(* IEC 61131-3 sources: RootPLC/conformance/cases/motion, 8 files *)

(* ---- ok_abort_and_relative.st ---- *)
(* spec: [motion.abort] [motion.move.relative]
   expect: ok
   libraries: RootMotion *)
TEST new_command_takes_control_without_a_jump
VAR
    ax : AXIS_REF;
    pw : MC_Power;
    m1 : MC_MoveAbsolute;
    m2 : MC_MoveRelative;
    i : INT;
    startPos : LREAL;
    vBefore : LREAL;
END_VAR
ax.CycleTime := 0.01;
pw(Enable := TRUE, Axis := ax);
FOR i := 1 TO 20 DO
    m1(Execute := TRUE, Position := 100.0, Velocity := 50.0, Acceleration := 100.0, Deceleration := 100.0, Axis := ax);
    RP_VirtualAxis(Axis := ax);
END_FOR;
startPos := ax.Position;
vBefore := ax.Velocity;
m2(Execute := TRUE, Distance := -5.0, Velocity := 50.0, Acceleration := 100.0, Deceleration := 100.0, Axis := ax);
m1(Execute := TRUE, Position := 100.0, Velocity := 50.0, Acceleration := 100.0, Deceleration := 100.0, Axis := ax);
ASSERT_TRUE(m1.CommandAborted);
ASSERT_FALSE(m1.Busy);
RP_VirtualAxis(Axis := ax);
ASSERT_TRUE(ABS(ax.Velocity - vBefore) <= 1.000001);
FOR i := 1 TO 300 DO
    m2(Execute := TRUE, Distance := -5.0, Velocity := 50.0, Acceleration := 100.0, Deceleration := 100.0, Axis := ax);
    RP_VirtualAxis(Axis := ax);
END_FOR;
ASSERT_TRUE(m2.Done);
ASSERT_TRUE(ABS(ax.Position - (startPos - 5.0)) < 0.000001);
END_TEST

(* ---- ok_errors_and_execute.st ---- *)
(* spec: [motion.errors] [motion.execute] [motion.power]
   expect: ok
   libraries: RootMotion *)
TEST command_on_unpowered_axis
VAR
    ax : AXIS_REF;
    mv : MC_MoveAbsolute;
END_VAR
mv(Execute := TRUE, Position := 10.0, Velocity := 5.0, Acceleration := 10.0, Deceleration := 10.0, Axis := ax);
ASSERT_TRUE(mv.Error);
ASSERT_EQ(UDINT#1, mv.ErrorID);
ASSERT_TRUE(ax.State = MC_AXIS_STATE#Disabled);
END_TEST

TEST invalid_parameter
VAR
    ax : AXIS_REF;
    pw : MC_Power;
    mv : MC_MoveAbsolute;
END_VAR
pw(Enable := TRUE, Axis := ax);
mv(Execute := TRUE, Position := 10.0, Velocity := 0.0, Acceleration := 10.0, Deceleration := 10.0, Axis := ax);
ASSERT_TRUE(mv.Error);
ASSERT_EQ(UDINT#3, mv.ErrorID);
ASSERT_TRUE(ax.State = MC_AXIS_STATE#Standstill);
END_TEST

TEST result_shows_one_call_after_execute_falls
VAR
    ax : AXIS_REF;
    pw : MC_Power;
    mv : MC_MoveAbsolute;
    i : INT;
END_VAR
ax.CycleTime := 0.1;
pw(Enable := TRUE, Axis := ax);
mv(Execute := TRUE, Position := 1.0, Velocity := 10.0, Acceleration := 100.0, Deceleration := 100.0, Axis := ax);
FOR i := 1 TO 20 DO
    mv(Execute := FALSE, Position := 1.0, Velocity := 10.0, Acceleration := 100.0, Deceleration := 100.0, Axis := ax);
    RP_VirtualAxis(Axis := ax);
    IF mv.Done THEN
        EXIT;
    END_IF;
END_FOR;
ASSERT_TRUE(mv.Done);
ASSERT_TRUE(ABS(ax.Position - 1.0) < 0.000001);
mv(Execute := FALSE, Position := 1.0, Velocity := 10.0, Acceleration := 100.0, Deceleration := 100.0, Axis := ax);
ASSERT_FALSE(mv.Done);
END_TEST

(* ---- ok_home.st ---- *)
(* spec: [motion.home] [motion.errors]
   expect: ok
   libraries: RootMotion *)
TEST home_sets_position
VAR
    ax : AXIS_REF;
    pw : MC_Power;
    hm : MC_Home;
END_VAR
hm(Execute := TRUE, Position := 0.0, Axis := ax);
ASSERT_TRUE(hm.Error);
ASSERT_EQ(UDINT#1, hm.ErrorID);
hm(Execute := FALSE, Position := 0.0, Axis := ax);
pw(Enable := TRUE, Axis := ax);
hm(Execute := TRUE, Position := 12.5, Axis := ax);
ASSERT_TRUE(hm.Done);
ASSERT_TRUE(ax.Homed);
ASSERT_TRUE(ABS(ax.Position - 12.5) < 0.000001);
ASSERT_TRUE(ax.State = MC_AXIS_STATE#Standstill);
END_TEST

(* ---- ok_limits_reset_stop.st ---- *)
(* spec: [motion.limits] [motion.reset] [motion.stop] [motion.errors]
   expect: ok
   libraries: RootMotion *)
TEST limit_error_reset_then_stop
VAR
    ax : AXIS_REF;
    pw : MC_Power;
    mvv : MC_MoveVelocity;
    mv : MC_MoveAbsolute;
    st : MC_Stop;
    rs : MC_Reset;
    i : INT;
END_VAR
ax.CycleTime := 0.01;
ax.LimitsEnabled := TRUE;
ax.PositiveLimit := 50.0;
ax.NegativeLimit := -50.0;
pw(Enable := TRUE, Axis := ax);
FOR i := 1 TO 600 DO
    mvv(Execute := TRUE, Velocity := 20.0, Acceleration := 100.0, Deceleration := 100.0, Axis := ax);
    RP_VirtualAxis(Axis := ax);
END_FOR;
mvv(Execute := TRUE, Velocity := 20.0, Acceleration := 100.0, Deceleration := 100.0, Axis := ax);
ASSERT_TRUE(ax.State = MC_AXIS_STATE#ErrorStop);
ASSERT_TRUE(mvv.Error);
ASSERT_EQ(UDINT#4, mvv.ErrorID);
ASSERT_TRUE(ABS(ax.Position - 50.0) < 0.000001);
ASSERT_TRUE(ABS(ax.Velocity) < 0.000001);
mv(Execute := TRUE, Position := 0.0, Velocity := 10.0, Acceleration := 100.0, Deceleration := 100.0, Axis := ax);
ASSERT_EQ(UDINT#2, mv.ErrorID);
rs(Execute := TRUE, Axis := ax);
ASSERT_TRUE(rs.Done);
ASSERT_TRUE(ax.State = MC_AXIS_STATE#Standstill);
ASSERT_EQ(UDINT#0, ax.ErrorID);
mvv(Execute := FALSE, Axis := ax);
mvv(Execute := FALSE, Axis := ax);
mvv(Execute := TRUE, Velocity := 10.0, Acceleration := 100.0, Deceleration := 100.0, Direction := MC_DIRECTION#Negative, Axis := ax);
RP_VirtualAxis(Axis := ax);
FOR i := 1 TO 50 DO
    st(Execute := TRUE, Deceleration := 100.0, Axis := ax);
    RP_VirtualAxis(Axis := ax);
END_FOR;
ASSERT_TRUE(st.Done);
ASSERT_TRUE(ax.State = MC_AXIS_STATE#Stopping);
mv(Execute := FALSE, Axis := ax);
mv(Execute := TRUE, Position := 0.0, Velocity := 10.0, Acceleration := 100.0, Deceleration := 100.0, Axis := ax);
ASSERT_EQ(UDINT#5, mv.ErrorID);
st(Execute := FALSE, Deceleration := 100.0, Axis := ax);
ASSERT_TRUE(ax.State = MC_AXIS_STATE#Standstill);
END_TEST

(* ---- ok_max_acceleration.st ---- *)
(* spec: [motion.axis] [motion.errors]
   expect: ok
   libraries: RootMotion *)
TEST command_above_machine_acceleration_is_rejected
VAR
    ax : AXIS_REF;
    pw : MC_Power;
    mv : MC_MoveAbsolute;
    hl : MC_Halt;
    i : INT;
END_VAR
ax.CycleTime := 0.01;
ax.MaxAcceleration := 500.0;
pw(Enable := TRUE, Axis := ax);
mv(Execute := TRUE, Position := 10.0, Velocity := 50.0, Acceleration := 600.0, Deceleration := 400.0, Axis := ax);
ASSERT_TRUE(mv.Error);
ASSERT_EQ(UDINT#3, mv.ErrorID);
ASSERT_TRUE(ax.State = MC_AXIS_STATE#Standstill);
mv(Execute := FALSE, Axis := ax);
FOR i := 1 TO 100 DO
    mv(Execute := TRUE, Position := 10.0, Velocity := 50.0, Acceleration := 500.0, Deceleration := 500.0, Axis := ax);
    RP_VirtualAxis(Axis := ax);
END_FOR;
ASSERT_TRUE(mv.Done);
hl(Execute := TRUE, Deceleration := 501.0, Axis := ax);
ASSERT_TRUE(hl.Error);
ASSERT_EQ(UDINT#3, hl.ErrorID);
END_TEST

(* ---- ok_move_absolute_profile.st ---- *)
(* spec: [motion.axis] [motion.cycle] [motion.power] [motion.profile] [motion.move.absolute] [motion.state]
   expect: ok
   libraries: RootMotion *)
(* 100 units at 50 units/s with 100 units/s2 both ways: 0.25 s + 2.0 s + 0.25 s
   = 2.5 s, so the goal is reached in cycle 250 and Done shows in cycle 251. *)
TEST trapezoid_reaches_target_on_time
VAR
    ax : AXIS_REF;
    pw : MC_Power;
    mv : MC_MoveAbsolute;
    i : INT;
    doneAt : INT := -1;
    vmax : LREAL;
    worstStep : LREAL;
    vPrev : LREAL;
END_VAR
ax.CycleTime := 0.01;
ASSERT_TRUE(ax.State = MC_AXIS_STATE#Disabled);
pw(Enable := TRUE, Axis := ax);
ASSERT_TRUE(pw.Status);
ASSERT_TRUE(ax.State = MC_AXIS_STATE#Standstill);
FOR i := 1 TO 400 DO
    mv(Execute := TRUE, Position := 100.0, Velocity := 50.0, Acceleration := 100.0, Deceleration := 100.0, Axis := ax);
    IF i = 1 THEN
        ASSERT_TRUE(ax.State = MC_AXIS_STATE#DiscreteMotion);
    END_IF;
    RP_VirtualAxis(Axis := ax);
    IF ax.Velocity > vmax THEN
        vmax := ax.Velocity;
    END_IF;
    IF ABS(ax.Velocity - vPrev) > worstStep THEN
        worstStep := ABS(ax.Velocity - vPrev);
    END_IF;
    vPrev := ax.Velocity;
    IF mv.Done AND doneAt < 0 THEN
        doneAt := i;
    END_IF;
END_FOR;
ASSERT_EQ(251, doneAt);
ASSERT_TRUE(ABS(ax.Position - 100.0) < 0.000001);
ASSERT_TRUE(ABS(vmax - 50.0) < 0.000001);
ASSERT_TRUE(worstStep <= 1.000001);
ASSERT_TRUE(ax.State = MC_AXIS_STATE#Standstill);
pw(Enable := FALSE, Axis := ax);
ASSERT_TRUE(ax.State = MC_AXIS_STATE#Disabled);
ASSERT_FALSE(pw.Status);
END_TEST

(* ---- ok_observe_axis_cycles.st ---- *)
(* spec: [motion.observe] [motion.cycle]
   expect: ok
   libraries: RootMotion *)
(* Reporting axis cycles to the toolchain changes nothing the program can
   see: the move behaves exactly as without the report. *)
TEST observed_move_is_unchanged
VAR
    ax : AXIS_REF;
    pw : MC_Power;
    mv : MC_MoveRelative;
    i : INT;
END_VAR
ax.CycleTime := 0.01;
pw(Enable := TRUE, Axis := ax);
FOR i := 1 TO 100 DO
    mv(Execute := TRUE, Distance := 10.0, Velocity := 50.0, Acceleration := 500.0, Deceleration := 500.0, Axis := ax);
    RP_VirtualAxis(Axis := ax);
END_FOR;
ASSERT_TRUE(mv.Done);
ASSERT_TRUE(ABS(ax.Position - 10.0) < 0.000001);
END_TEST

(* ---- ok_velocity_halt_read.st ---- *)
(* spec: [motion.move.velocity] [motion.halt] [motion.read] [motion.state]
   expect: ok
   libraries: RootMotion *)
TEST velocity_then_halt
VAR
    ax : AXIS_REF;
    pw : MC_Power;
    mvv : MC_MoveVelocity;
    hl : MC_Halt;
    rd : MC_ReadStatus;
    rp : MC_ReadActualPosition;
    i : INT;
END_VAR
ax.CycleTime := 0.01;
pw(Enable := TRUE, Axis := ax);
FOR i := 1 TO 100 DO
    mvv(Execute := TRUE, Velocity := 20.0, Acceleration := 100.0, Deceleration := 100.0, Direction := MC_DIRECTION#Negative, Axis := ax);
    RP_VirtualAxis(Axis := ax);
END_FOR;
mvv(Execute := TRUE, Velocity := 20.0, Acceleration := 100.0, Deceleration := 100.0, Direction := MC_DIRECTION#Negative, Axis := ax);
ASSERT_TRUE(mvv.InVelocity);
ASSERT_TRUE(ABS(ax.Velocity + 20.0) < 0.000001);
rd(Enable := TRUE, Axis := ax);
ASSERT_TRUE(rd.ContinuousMotion);
ASSERT_FALSE(rd.Standstill);
rp(Enable := TRUE, Axis := ax);
ASSERT_TRUE(rp.Valid);
ASSERT_TRUE(ABS(rp.Position - ax.Position) < 0.000001);
FOR i := 1 TO 50 DO
    hl(Execute := TRUE, Deceleration := 100.0, Axis := ax);
    mvv(Execute := TRUE, Velocity := 20.0, Acceleration := 100.0, Deceleration := 100.0, Direction := MC_DIRECTION#Negative, Axis := ax);
    RP_VirtualAxis(Axis := ax);
END_FOR;
ASSERT_TRUE(hl.Done);
ASSERT_TRUE(mvv.CommandAborted);
ASSERT_FALSE(mvv.InVelocity);
ASSERT_TRUE(ax.State = MC_AXIS_STATE#Standstill);
rd(Enable := TRUE, Axis := ax);
ASSERT_TRUE(rd.Standstill);
END_TEST
